(* IEC 61131-3 sources: sis-interlock-demo/src/POUs/Sis/F_SisBitMask, 2 files *)

(* ---- F_SisBitMask.decl.st ---- *)
// Назначение: маска одного бита по индексу с единицы: SHL(WORD_BIT0, uiIdx − 1); вне 1..16 — 0.
// Автор:      kr0nsch
// Версия:     0.1.0
// Документ:   docs/DESIGN.md, раздел «8.2 Функции работы с битами»
// ВНИМАНИЕ:   код демонстрационный и не предназначен для систем безопасности. Реальная ПАЗ
//             требует определения SIL, сертифицированных аппаратных и программных средств
//             и валидации по ГОСТ Р МЭК 61511.
FUNCTION F_SisBitMask : WORD
VAR_INPUT
    uiIdx : UINT;    // индекс причины или следствия, 1..16
END_VAR

(* ---- F_SisBitMask.impl.st ---- *)
IF uiIdx >= 1 AND uiIdx <= GVL_Const.WORD_BITS THEN
    F_SisBitMask := SHL(GVL_Const.WORD_BIT0, uiIdx - 1);
ELSE
    F_SisBitMask := 0;
END_IF
